// TIA Portal V20 export
// export: Created 2026-10-20T12:41:00.7160763Z, ExportSetting WithDefaults, DisplayName Totally Integrated Automation Portal, DisplayVersion V20 Update 6, DisplayName TIA Portal Openness, DisplayVersion V20 Update 6, DisplayName TIA Portal Version Control Interface, DisplayVersion V20 Update 6, DisplayName SINAMICS Startdrive Advanced, DisplayVersion V20 SP1, DisplayName SINAMICS Startdrive G130, G150, S120, S150, SINAMICS MV, G220, S200, S210, DisplayVersion V20 SP1, DisplayName SINAMICS Startdrive G110M, G120, G120C, G120D, G120P, G115D, DisplayVersion V20 SP1, DisplayName STEP 7 Professional, DisplayVersion V20 Update 6, DisplayName STEP 7 Safety, DisplayVersion V20 Update 2, DisplayName WinCC Basic/Comfort/Advanced, DisplayVersion V20 Update 6, DisplayName WinCC Unified, DisplayVersion V20 Update 6
DATA_BLOCK "SICK_Lector_Control_DB_4"   // DB153
VERSION : 0.1
// stored: AutoNumber true, DBAccessibleFromOPCUA true, InstanceOfName SICK_Lector_Control_FB, InstanceOfType FB
"SICK_Lector_Control_FB"
   // VAR_INPUT
   //    Rd_Done : Bool;
   //    Req_Done : Bool;
   //    Req_Busy : Bool;
   //    Error : Bool;
   //    arrResult : Array[1..200] of Byte;
   //    iCounter : USInt;
   //    iLength : Int;
   //    Error_Code : DWord;
   // END_VAR
   // VAR_OUTPUT
   //    Test_Comm : Bool;
   //    Enable_Trigger : Bool;
   //    Disable_Trigger : Bool;
   //    Enable_Req : Bool;
   //    Result : String;
   //    Test_OK : Bool;
   // END_VAR
   // VAR_IN_OUT
   //    Test_Comm_HMI : Bool;
   //    Enable_HMI : Bool;
   //    Disable_HMI : Bool;
   //    Auto_Start_Lector : Bool;
   //    Auto_Stop_Lector : Bool;
   // END_VAR
   // VAR
   //    "Timer" { S7_SetPoint := 'True'} : TON_TIME;
   //    R_Done_DB { S7_SetPoint := 'True'} : R_TRIG;
   //    T_Reset_DB { S7_SetPoint := 'True'} : TON_TIME;
   // END_VAR
BEGIN
END_DATA_BLOCK
